// TIA Portal V20 export
Screen "SafetyZone05Overview"  1276x673
  ScreenItem "Button_Overview_LegendᆉY2" at 1185,2 size 90x60  Type=HmiButton
  ScreenItem "Button_Back" at 2,4 size 90x60  Type=HmiButton
  ScreenItem "Rectangle_12" at 662,625 size 482x8  Type=HmiRectangle
  ScreenItem "Line_Header_X0_Y64" at -11,64 size 1280x0  Type=HmiLine
  ScreenItem "文本域_16" at 31,683 size 50x20  Type=HmiTextBox
  ScreenItem "Emerg_4" at 28,696 size 52x56  Type=HmiSymbolicIOField
  ScreenItem "Graphic view_15" at 32,276 size 46x35  Type=HmiGraphicView
  ScreenItem "Graphic view_19" at 1199,284 size 46x35  Type=HmiGraphicView
  ScreenItem "Faceplate container_15" at 862,527 size 152x87  Type=HmiFaceplateContainer
  ScreenItem "Faceplate container_21" at 472,389 size 110x139  Type=HmiFaceplateContainer
  ScreenItem "Faceplate container_6" at 735,470 size 110x138  Type=HmiFaceplateContainer
  ScreenItem "Rectangle_5" at 18,77 size 549x8  Type=HmiRectangle
  ScreenItem "Rectangle_6" at 745,77 size 513x8  Type=HmiRectangle
  ScreenItem "Rectangle_7" at 1174,154 size 160x8  Type=HmiRectangle
  ScreenItem "Rectangle_11" at 1112,487 size 284x8  Type=HmiRectangle
  ScreenItem "Rectangle_13" at 16,625 size 648x8  Type=HmiRectangle
  ScreenItem "Rectangle_14" at -60,152 size 160x8  Type=HmiRectangle
  ScreenItem "Rectangle_15" at 146,566 size 109x8  Type=HmiRectangle
  ScreenItem "Graphic view_4" at 449,279 size 46x35  Type=HmiGraphicView
  ScreenItem "图形 IO 域_26" at 13,234 size 15x122  Type=HmiSymbolicIOField
  ScreenItem "图形 IO 域_15" at 1247,238 size 15x122  Type=HmiSymbolicIOField
  ScreenItem "Button_Overview_LegendᆉY2_1" at 1092,2 size 90x60  Type=HmiButton
  ScreenItem "矩形_1" at 1146,625 size 14x11  Type=HmiRectangle
  ScreenItem "线_1" at 1159,640 size 47x13  Type=HmiLine
  ScreenItem "矩形_2" at 1159,625 size 48x11  Type=HmiRectangle
  ScreenItem "矩形_3" at 1206,625 size 14x11  Type=HmiRectangle
  ScreenItem "Rectangle_30" at 1220,627 size 36x8  Type=HmiRectangle
  ScreenItem "Title_ScreenOverview_X390_Y2_1" at 384,4 size 510x57  Type=HmiTextBox
  ScreenItem "矩形_4" at 565,76 size 14x11  Type=HmiRectangle
  ScreenItem "线_2" at 578,91 size 47x13  Type=HmiLine
  ScreenItem "矩形_5" at 578,76 size 48x11  Type=HmiRectangle
  ScreenItem "矩形_6" at 625,76 size 14x11  Type=HmiRectangle
  ScreenItem "Rectangle_2" at 639,77 size 106x8  Type=HmiRectangle
  ScreenItem "Rectangle_3" at 24,373 size 565x8  Type=HmiRectangle
  ScreenItem "Rectangle_4" at 465,495 size 257x8  Type=HmiRectangle
  ScreenItem "Faceplate container_26" at 601,376 size 152x87  Type=HmiFaceplateContainer
  ScreenItem "Graphic view_3" at 691,270 size 46x35  Type=HmiGraphicView
  ScreenItem "Rectangle_8" at 437,143 size 142x8  Type=HmiRectangle
  ScreenItem "Faceplate container_3" at 843,232 size 362x136  Type=HmiFaceplateContainer
  ScreenItem "Faceplate container_1" at 855,90 size 110x140  Type=HmiFaceplateContainer
  ScreenItem "Faceplate container_4" at 1094,90 size 110x140  Type=HmiFaceplateContainer
  ScreenItem "Faceplate container_5" at 1094,367 size 110x140  Type=HmiFaceplateContainer
  ScreenItem "Faceplate container_7" at 38,527 size 152x87  Type=HmiFaceplateContainer
  ScreenItem "Faceplate container_8" at 214,527 size 152x87  Type=HmiFaceplateContainer
  ScreenItem "Faceplate container_9" at 437,534 size 152x87  Type=HmiFaceplateContainer
  ScreenItem "Faceplate container_16" at 664,92 size 152x87  Type=HmiFaceplateContainer
  ScreenItem "Faceplate container_10" at 973,367 size 110x140  Type=HmiFaceplateContainer
  ScreenItem "Faceplate container_2" at 973,90 size 110x140  Type=HmiFaceplateContainer
  ScreenItem "Faceplate container_11" at 855,367 size 110x140  Type=HmiFaceplateContainer
  ScreenItem "Faceplate container_12" at 612,467 size 100x138  Type=HmiFaceplateContainer
  ScreenItem "Faceplate container_13" at 71,230 size 362x136  Type=HmiFaceplateContainer
  ScreenItem "Rectangle_1" at -116,492 size 277x8  Type=HmiRectangle
  ScreenItem "Rectangle_9" at 32,515 size 352x8  Type=HmiRectangle
  ScreenItem "Rectangle_10" at 334,570 size 100x8  Type=HmiRectangle
  ScreenItem "Faceplate container_14" at 196,90 size 152x87  Type=HmiFaceplateContainer
  ScreenItem "Emerg_1" at 521,77 size 52x56  Type=HmiSymbolicIOField
  ScreenItem "文本域_1" at 518,130 size 58x19  Type=HmiTextBox
  ScreenItem "Emerg_2" at 1092,577 size 52x56  Type=HmiSymbolicIOField
  ScreenItem "文本域_2" at 1089,563 size 58x19  Type=HmiTextBox
